// TIA Portal V21 export
// export: Created 2026-11-08T21:35:34.1352715Z, ExportSetting WithDefaults, DisplayName Totally Integrated Automation Portal, DisplayVersion V21 Update 3, DisplayName STEP 7 Professional, DisplayVersion V21 Update 3, DisplayName STEP 7 Safety, DisplayVersion V21, DisplayName Tech WebApplication, DisplayVersion V21, DisplayName WinCC Basic/Comfort/Advanced, DisplayVersion V21 Update 3, DisplayName WinCC Unified, DisplayVersion V21 Update 3
FUNCTION_BLOCK "FB_StlC_037"   // FB86, STL
TITLE = STL call ReadFromArrayDB
{ S7_Optimized_Access := 'TRUE' }
VERSION : 0.1
// stored: AutoNumber true, IsRetainMemResEnabled false, MemoryReserve 100, UDAEnableTagReadback false
   VAR_INPUT
      di1 : DInt;
   END_VAR
   VAR_OUTPUT
      io : Int;
   END_VAR
   VAR
      val : Int;
   END_VAR
BEGIN

NETWORK
TITLE = 037 ReadFromArrayDB
      CALL  ReadFromArrayDB
      ( db      := "ArrDB",
        index   := #di1,
        Ret_Val := #io,
        value   := #val
      );

NETWORK
TITLE = 038 WriteToArrayDB
      CALL  WriteToArrayDB
      ( db      := "ArrDB",
        index   := #di1,
        value   := #val,
        Ret_Val := #io
      );
END_FUNCTION_BLOCK
